FUNCTION_BLOCK basicValvulaCoester (* Logica do atuador Coester CSR (Modbus TCP) *)
  (* Standard: 61499-2 *)
  (* Version 2.5, 12/11/2026, Hidryco, Hidryco, 2.5: mapa revisado pelo MN_065 rev.3 (Modbus RTU, painel BLE): leitura 101-109 e comandos conferidos; posicao (word 105) = bits 0-7 parte inteira, bits 8-15 parte decimal - usa so o byte baixo, sem filtro de faixa (antes a word inteira dava valores acima de 1000). 2.4: posicao (Word 5) so atualiza com leitura de 0 a 100; fora da faixa mantem a ultima valida (antes era limitada, e um valor acima de 1000 virava 100 %%). 2.3: falha do atuador (alarmes da comunicacao) nao bloqueia o comando (fica disponivel em automatico) e nao muda a cor (sem animacao de falha); continua no alarme, no STS_ALARME e no diagnostico. 2.2: stsAlarme para a IO List da Nereda. 2.1: leituras 100 a 108 (posicao, torque, temperatura, tempo de percurso, status 2, alarmes), falha do atuador, posicionar por comando e parar so com cfgPosicionador (Word 2 de escrita). 2.0: refeito simples. *)
  PACKAGE Hidryco.HidrycoLib;
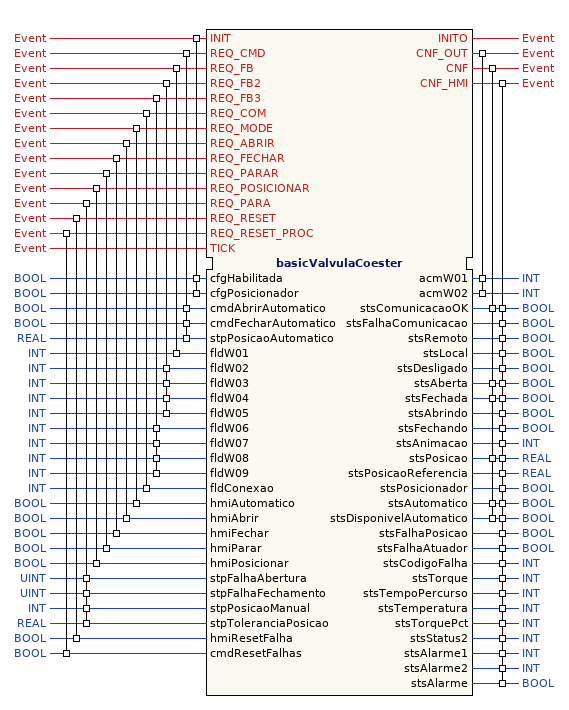
  EVENT_INPUT
    INIT WITH cfgHabilitada, cfgPosicionador; (* Inicializacao *)
    REQ_CMD WITH cmdAbrirAutomatico, cmdFecharAutomatico, stpPosicaoAutomatico; (* Processo: comandos do automatico *)
    REQ_FB WITH fldW01; (* Leitura Modbus: status 1 (endereco 100) *)
    REQ_FB2 WITH fldW02, fldW03, fldW04, fldW05; (* Leitura Modbus: enderecos 101 a 104 *)
    REQ_FB3 WITH fldW06, fldW07, fldW08, fldW09; (* Leitura Modbus: enderecos 105 a 108 *)
    REQ_COM WITH fldConexao; (* Status da conexao Modbus (connStatusInt) *)
    REQ_MODE WITH hmiAutomatico; (* IHM: modo *)
    REQ_ABRIR WITH hmiAbrir; (* IHM: abrir (manual) *)
    REQ_FECHAR WITH hmiFechar; (* IHM: fechar (manual) *)
    REQ_PARAR WITH hmiParar; (* IHM: parar (manual, so posicionador) *)
    REQ_POSICIONAR WITH hmiPosicionar; (* IHM: posicionar (manual, so posicionador) *)
    REQ_PARA WITH stpFalhaAbertura, stpFalhaFechamento, stpPosicaoManual, stpToleranciaPosicao; (* IHM: parametros *)
    REQ_RESET WITH hmiResetFalha; (* IHM: reset *)
    REQ_RESET_PROC WITH cmdResetFalhas; (* Processo: reset *)
    TICK; (* Base de tempo de 1 s *)
  END_EVENT
  EVENT_OUTPUT
    INITO; (* Inicializacao concluida *)
    CNF_OUT WITH acmW01, acmW02; (* Escrita Modbus (comando e posicao) *)
    CNF WITH stsDisponivelAutomatico, stsAberta, stsFechada, stsPosicao, stsAutomatico, stsComunicacaoOK; (* Status para o processo (na mudanca) *)
    CNF_HMI WITH stsComunicacaoOK, stsFalhaComunicacao, stsRemoto, stsLocal, stsDesligado, stsAberta, stsFechada, stsAbrindo, stsFechando, stsAnimacao, stsAutomatico, stsDisponivelAutomatico, stsFalhaPosicao, stsPosicionador, stsPosicao, stsPosicaoReferencia, stsFalhaAtuador, stsCodigoFalha, stsTorque, stsTempoPercurso, stsTemperatura, stsTorquePct, stsStatus2, stsAlarme1, stsAlarme2, stsAlarme; (* Status para a IHM (1 s e no comando) *)
  END_EVENT
  VAR_INPUT
    cfgHabilitada : BOOL := TRUE; (* FALSE = equipamento futuro: sem comunicacao esperada, sem alarme, fora do automatico *)
    cfgPosicionador : BOOL := FALSE; (* TRUE = posicionar e parar (700-VC-01); FALSE = so abrir e fechar *)
    cmdAbrirAutomatico : BOOL; (* Automatico: abrir *)
    cmdFecharAutomatico : BOOL; (* Automatico: fechar *)
    stpPosicaoAutomatico : REAL; (* Automatico: posicao desejada (%) - so posicionador *)
    fldW01 : INT; (* Word 1: status 1 (b0 local, b1 remoto, b2 desligado, b3 aberta, b4 fechada, b6 abrindo, b7 fechando) *)
    fldW02 : INT; (* Word 2: status 2 *)
    fldW03 : INT; (* Word 3: alarmes 1 *)
    fldW04 : INT; (* Word 4: alarmes 2 *)
    fldW05 : INT; (* Word 5: posicao (%) *)
    fldW06 : INT; (* Word 6: torque (Nm) *)
    fldW07 : INT; (* Word 7: tempo de percurso (s) *)
    fldW08 : INT; (* Word 8: temperatura (valor - 19 = graus C) *)
    fldW09 : INT; (* Word 9: torque (%) *)
    fldConexao : INT; (* Conexao Modbus: 1 = online *)
    hmiAutomatico : BOOL; (* IHM: TRUE = automatico *)
    hmiAbrir : BOOL; (* IHM: abrir *)
    hmiFechar : BOOL; (* IHM: fechar *)
    hmiParar : BOOL; (* IHM: parar *)
    hmiPosicionar : BOOL; (* IHM: posicionar *)
    stpFalhaAbertura : UINT; (* Tempo maximo para abrir (s); 0 = sem supervisao *)
    stpFalhaFechamento : UINT; (* Tempo maximo para fechar (s); 0 = sem supervisao *)
    stpPosicaoManual : INT; (* Posicao desejada em manual (%) *)
    stpToleranciaPosicao : REAL; (* Tolerancia da posicao (%); 0 = 2 % *)
    hmiResetFalha : BOOL; (* IHM: reset *)
    cmdResetFalhas : BOOL; (* Processo: reset (vale com TRUE) *)
  END_VAR
  VAR_OUTPUT
    acmW01 : INT; (* Word 1 de escrita (endereco 0): pulso b0 abrir, b1 fechar, b2 parar, b4 posicionar, b8 quitar alarmes *)
    acmW02 : INT; (* Word 2 de escrita (endereco 1): posicao desejada 0-100 % (so posicionador) *)
    stsComunicacaoOK : BOOL; (* Comunicacao OK *)
    stsFalhaComunicacao : BOOL; (* Falha de comunicacao *)
    stsRemoto : BOOL; (* Seletor em remoto *)
    stsLocal : BOOL; (* Seletor em local *)
    stsDesligado : BOOL; (* Seletor em desligado *)
    stsAberta : BOOL; (* Aberta *)
    stsFechada : BOOL; (* Fechada *)
    stsAbrindo : BOOL; (* Abrindo *)
    stsFechando : BOOL; (* Fechando *)
    stsAnimacao : INT; (* 0 fechada, 1 aberta, 2 falha, 3 intermediaria parada, 4 abrindo, 5 fechando *)
    stsPosicao : REAL; (* Posicao real (%) - Word 5 *)
    stsPosicaoReferencia : REAL; (* Ultima posicao enviada (%) *)
    stsPosicionador : BOOL; (* Copia de cfgPosicionador para a IHM *)
    stsAutomatico : BOOL; (* Modo automatico *)
    stsDisponivelAutomatico : BOOL; (* Pode ser comandada pelo automatico *)
    stsFalhaPosicao : BOOL; (* Nao abriu / nao fechou / nao posicionou no tempo (memorizada ate o reset) *)
    stsFalhaAtuador : BOOL; (* Falha do atuador (memorizada ate o reset) *)
    stsCodigoFalha : INT; (* Codigo da falha do atuador *)
    stsTorque : INT; (* Torque (Nm) *)
    stsTempoPercurso : INT; (* Tempo de percurso (s) *)
    stsTemperatura : INT; (* Temperatura (graus C) *)
    stsTorquePct : INT; (* Torque (%) *)
    stsStatus2 : INT; (* Word 2 *)
    stsAlarme1 : INT; (* Word 3 *)
    stsAlarme2 : INT; (* Word 4 *)
    stsAlarme : BOOL; (* Alarme: falha de comunicacao OU falha do atuador OU nao abriu/fechou/posicionou *)
  END_VAR
  VAR
    initDone : BOOL;
    comRecebido : BOOL;
    bComOk : BOOL;
    w01 : WORD;
    w02 : WORD;
    w03 : WORD;
    w04 : WORD;
    bFalhaAtiva : BOOL;
    codAtivo : INT;
    bAuto : BOOL := TRUE;
    bCmdMan : INT;
    bSpMan : REAL;
    bForca : BOOL;
    bPode : BOOL;
    bAlvo : INT;
    bAlvoAnt : INT := -1;
    bSp : REAL;
    bSpEnviado : REAL;
    bSubindo : BOOL;
    cBanda : REAL := 2.0;
    rTol : REAL;
    tLim : DINT;
    wPulso : WORD;
    tPulso : INT;
    cTempoPulso : INT := 2;
    wCmd : WORD;
    tReset : INT;
    tPos : INT;
    oldW01 : INT := -1;
    oldW02 : INT := -1;
    oldProc : INT := -1;
    oldPos : REAL := -1.0;
    nProc : INT;
    primeiro : BOOL := TRUE;
  END_VAR
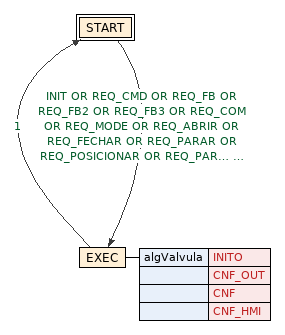
  EC_STATES
    START; (* Estado inicial *)
    EXEC : algValvula -> INITO, -> CNF_OUT, -> CNF, -> CNF_HMI; (* Executa a logica; o algoritmo decide quais eventos saem *)
  END_STATES
  EC_TRANSITIONS
    START TO EXEC := INIT OR REQ_CMD OR REQ_FB OR REQ_FB2 OR REQ_FB3 OR REQ_COM OR REQ_MODE OR REQ_ABRIR OR REQ_FECHAR OR REQ_PARAR OR REQ_POSICIONAR OR REQ_PARA OR REQ_RESET OR REQ_RESET_PROC OR TICK;
    EXEC TO START := 1;
  END_TRANSITIONS
  ALGORITHM algValvula IN ST: (* Logica completa da valvula (um unico algoritmo) *)
(* =====================================================================
   basicValvulaCoester 2.1 - logica do CAT Atuador_Coester (HidrycoLib)
   Atuador Coester CSR por Modbus TCP (mapa medido em campo):
   - leitura 100..108 = Words 1 a 9: status 1, status 2, alarmes 1 e 2,
     posicao (%), torque (Nm), tempo de percurso (s), temperatura (-19),
     torque (%);
   - escrita 0..1: Word 1 = comando EM PULSO de cTempoPulso s (b0 abrir,
     b1 fechar, b2 parar, b4 posicionar, b8 quitar alarmes); Word 2 =
     posicao desejada 0-100 %. O atuador retem o comando (MN_058 4.2.22);
     posicionar e "por comando" (padrao, MN_058 4.2.11): grava a Word 2 e
     pulsa o b4.
   - cfgPosicionador = TRUE (700-VC-01): posicionar e parar; no automatico
     segue stpPosicaoAutomatico e reposiciona quando ela muda cBanda (2 %)
     ou mais. FALSE: so abrir e fechar.
   - so comanda em remoto e com comunicacao OK; voltar a remoto repete o
     comando vigente; em manual cada botao repete o pulso;
   - "nao abriu / nao fechou / nao posicionou": o fim de curso (ou a
     posicao, com a tolerancia) nao veio no tempo configurado (0 = sem
     supervisao); memoriza ate o reset e pulsa parar;
   - falha do atuador: status 2 b0-b2, alarme 1 b1-b12, alarme 2 b0, b1,
     b4-b8; memoriza ate o reset; so informa (alarme e diagnostico):
     nao bloqueia o comando nem muda a cor da valvula;
   - cfgHabilitada = FALSE (equipamento futuro): sem alarme, fora do automatico.
   ===================================================================== *)

INITO   := FALSE;
CNF_OUT := FALSE;
CNF     := FALSE;
CNF_HMI := FALSE;

IF REQ_COM THEN
    comRecebido := TRUE;
END_IF;
IF INIT THEN
    initDone := TRUE;
    INITO    := TRUE;
END_IF;
IF NOT initDone THEN
    RETURN;
END_IF;

(* ---- 1. Leituras ---- *)
bComOk := cfgHabilitada AND comRecebido AND (fldConexao = 1);
w01 := INT_TO_WORD(fldW01);
w02 := INT_TO_WORD(fldW02);
w03 := INT_TO_WORD(fldW03);
w04 := INT_TO_WORD(fldW04);
IF bComOk THEN
    stsLocal     := (w01 AND 16#0001) <> 16#0000;
    stsRemoto    := (w01 AND 16#0002) <> 16#0000;
    stsDesligado := (w01 AND 16#0004) <> 16#0000;
    stsAberta    := (w01 AND 16#0008) <> 16#0000;
    stsFechada   := (w01 AND 16#0010) <> 16#0000;
    stsAbrindo   := (w01 AND 16#0040) <> 16#0000;
    stsFechando  := (w01 AND 16#0080) <> 16#0000;
    (* posicao (MN_065 rev.3, painel BLE, word 105): bits 0-7 = parte inteira (%), bits 8-15 = parte
       decimal; usa so o byte baixo (parte inteira) *)
    stsPosicao := INT_TO_REAL(WORD_TO_INT(INT_TO_WORD(fldW05) AND 16#00FF));
    stsTorque        := fldW06;
    stsTempoPercurso := fldW07;
    stsTemperatura   := fldW08 - 19;
    stsTorquePct     := fldW09;
    stsStatus2       := fldW02;
    stsAlarme1       := fldW03;
    stsAlarme2       := fldW04;
    bFalhaAtiva := ((w02 AND 16#0007) <> 16#0000) OR ((w03 AND 16#1FFE) <> 16#0000) OR ((w04 AND 16#01F3) <> 16#0000);
ELSE
    stsLocal := FALSE; stsRemoto := FALSE; stsDesligado := FALSE;
    stsAberta := FALSE; stsFechada := FALSE; stsAbrindo := FALSE; stsFechando := FALSE;
    bFalhaAtiva := FALSE;                      (* posicao e medicoes ficam no ultimo valor lido *)
END_IF;
stsComunicacaoOK    := bComOk;
stsFalhaComunicacao := cfgHabilitada AND NOT bComOk;
stsPosicionador     := cfgPosicionador;

(* codigo da falha ativa de maior prioridade (texto na IHM) *)
codAtivo := 0;
IF bFalhaAtiva THEN
    IF ((w02 AND 16#0001) <> 16#0000) OR ((w03 AND 16#0800) <> 16#0000) THEN codAtivo := 1;      (* falta de fase *)
    ELSIF ((w02 AND 16#0002) <> 16#0000) OR ((w03 AND 16#0040) <> 16#0000) THEN codAtivo := 2;   (* sobreaquecimento *)
    ELSIF ((w02 AND 16#0004) <> 16#0000) OR ((w03 AND 16#1000) <> 16#0000) THEN codAtivo := 3;   (* sem programacao *)
    ELSIF (w03 AND 16#0002) <> 16#0000 THEN codAtivo := 4;   (* parada local de emergencia *)
    ELSIF (w03 AND 16#0004) <> 16#0000 THEN codAtivo := 5;   (* torque na abertura *)
    ELSIF (w03 AND 16#0008) <> 16#0000 THEN codAtivo := 6;   (* torque no fechamento *)
    ELSIF (w03 AND 16#0010) <> 16#0000 THEN codAtivo := 7;   (* travado *)
    ELSIF (w03 AND 16#0020) <> 16#0000 THEN codAtivo := 8;   (* operacao incompleta *)
    ELSIF (w03 AND 16#0080) <> 16#0000 THEN codAtivo := 9;   (* falha ao energizar o motor *)
    ELSIF (w03 AND 16#0100) <> 16#0000 THEN codAtivo := 10;  (* motor energizado apos fim de curso *)
    ELSIF (w03 AND 16#0200) <> 16#0000 THEN codAtivo := 11;  (* motor energizado apos parada *)
    ELSIF (w03 AND 16#0400) <> 16#0000 THEN codAtivo := 12;  (* falha de comando *)
    ELSIF (w04 AND 16#0001) <> 16#0000 THEN codAtivo := 13;  (* tensao alta *)
    ELSIF (w04 AND 16#0002) <> 16#0000 THEN codAtivo := 14;  (* tensao baixa *)
    ELSIF (w04 AND 16#0030) <> 16#0000 THEN codAtivo := 15;  (* fim de curso mecanico ultrapassado *)
    ELSIF (w04 AND 16#00C0) <> 16#0000 THEN codAtivo := 16;  (* fim de curso programado ultrapassado *)
    ELSIF (w04 AND 16#0100) <> 16#0000 THEN codAtivo := 17;  (* cartao de rede nao detectado *)
    END_IF;
    stsFalhaAtuador := TRUE;                   (* memoriza ate o reset *)
    stsCodigoFalha  := codAtivo;
END_IF;

(* ---- 2. Reset (IHM ou processo) ---- *)
IF (REQ_RESET AND hmiResetFalha) OR (REQ_RESET_PROC AND cmdResetFalhas) THEN
    stsFalhaAtuador := bFalhaAtiva;            (* continua se a falha ainda esta ativa no atuador *)
    IF NOT bFalhaAtiva THEN
        stsCodigoFalha := 0;
    END_IF;
    stsFalhaPosicao := FALSE;
    tPos   := 0;
    tReset := 3;                               (* quitar alarmes no atuador por 3 s *)
END_IF;
IF TICK AND (tReset > 0) THEN
    tReset := tReset - 1;
END_IF;

(* ---- 3. Modo, parametros e comandos manuais ---- *)
IF REQ_MODE THEN
    bAuto := hmiAutomatico;
    bCmdMan := 0;                              (* troca de modo: nenhum comando manual *)
END_IF;
IF stpToleranciaPosicao > 0.0 THEN
    rTol := stpToleranciaPosicao;
ELSE
    rTol := 2.0;
END_IF;
bForca := FALSE;
IF NOT bAuto THEN
    IF REQ_ABRIR AND hmiAbrir THEN bCmdMan := 1; bForca := TRUE; END_IF;
    IF REQ_FECHAR AND hmiFechar THEN bCmdMan := 2; bForca := TRUE; END_IF;
    IF cfgPosicionador THEN
        IF REQ_PARAR AND hmiParar THEN bCmdMan := 4; bForca := TRUE; END_IF;
        IF REQ_POSICIONAR AND hmiPosicionar THEN
            bCmdMan := 3; bForca := TRUE;
            bSpMan := LIMIT(0.0, INT_TO_REAL(stpPosicaoManual), 100.0);
        END_IF;
    END_IF;
END_IF;

(* ---- 4. Comando desejado: 0 nenhum, 1 abrir, 2 fechar, 3 posicionar, 4 parar ---- *)
bPode := bComOk AND stsRemoto;
bSp := bSpEnviado;
IF NOT bPode THEN
    bAlvo := 0;                                (* fora de remoto ou sem comunicacao: nao comanda *)
ELSIF stsFalhaPosicao THEN
    bAlvo := 4;                                (* nao abriu / nao fechou / nao posicionou: para *)
ELSIF bAuto THEN
    IF cfgPosicionador THEN
        bAlvo := 3;
        bSp := LIMIT(0.0, stpPosicaoAutomatico, 100.0);
    ELSIF cmdAbrirAutomatico AND NOT cmdFecharAutomatico THEN
        bAlvo := 1;
    ELSIF cmdFecharAutomatico AND NOT cmdAbrirAutomatico THEN
        bAlvo := 2;
    ELSE
        bAlvo := 0;
    END_IF;
ELSE
    bAlvo := bCmdMan;
    IF bCmdMan = 3 THEN
        bSp := bSpMan;
    END_IF;
END_IF;

(* ---- 5. Pulso de comando ---- *)
IF TICK AND (tPulso > 0) THEN
    tPulso := tPulso - 1;
END_IF;
IF (bAlvo <> bAlvoAnt) OR (bForca AND bPode) OR ((bAlvo = 3) AND (ABS(bSp - bSpEnviado) >= cBanda)) THEN
    CASE bAlvo OF
        1: wPulso := 16#0001;
        2: wPulso := 16#0002;
        3: wPulso := 16#0010;
        4: wPulso := 16#0004;
    ELSE
        wPulso := 16#0000;
    END_CASE;
    IF bAlvo = 3 THEN
        bSubindo   := bSp >= stsPosicao;
        bSpEnviado := bSp;
    ELSIF bAlvo = 1 THEN
        bSpEnviado := 100.0;
    ELSIF bAlvo = 2 THEN
        bSpEnviado := 0.0;
    END_IF;
    IF wPulso <> 16#0000 THEN
        tPulso := cTempoPulso;
    ELSE
        tPulso := 0;
    END_IF;
    bAlvoAnt := bAlvo;
    tPos := 0;
END_IF;
IF tPulso > 0 THEN
    wCmd := wPulso;
ELSE
    wCmd := 16#0000;
END_IF;
IF tReset > 0 THEN
    wCmd := wCmd OR 16#0100;
END_IF;
acmW01 := WORD_TO_INT(wCmd);
acmW02 := REAL_TO_INT(LIMIT(0.0, bSpEnviado, 100.0));
stsPosicaoReferencia := bSpEnviado;
IF (acmW01 <> oldW01) OR (acmW02 <> oldW02) OR TICK OR primeiro THEN
    CNF_OUT := TRUE;
    oldW01 := acmW01;
    oldW02 := acmW02;
END_IF;

(* ---- 6. Nao abriu / nao fechou / nao posicionou ---- *)
IF TICK THEN
    tLim := 0;
    IF bPode THEN
        IF (bAlvo = 1) AND NOT stsAberta THEN
            tLim := UINT_TO_DINT(stpFalhaAbertura);
        ELSIF (bAlvo = 2) AND NOT stsFechada THEN
            tLim := UINT_TO_DINT(stpFalhaFechamento);
        ELSIF (bAlvo = 3) AND (ABS(stsPosicao - bSpEnviado) > rTol) THEN
            IF bSubindo THEN
                tLim := UINT_TO_DINT(stpFalhaAbertura);
            ELSE
                tLim := UINT_TO_DINT(stpFalhaFechamento);
            END_IF;
        END_IF;
    END_IF;
    IF tLim > 0 THEN
        tPos := tPos + 1;
        IF INT_TO_DINT(tPos) >= tLim THEN
            stsFalhaPosicao := TRUE;
        END_IF;
    ELSE
        tPos := 0;
    END_IF;
END_IF;

(* ---- 7. Saidas ---- *)
stsAutomatico := bAuto;
stsDisponivelAutomatico := bComOk AND stsRemoto AND bAuto AND NOT stsFalhaPosicao;   (* falha do atuador nao bloqueia *)
IF NOT bComOk OR stsFalhaPosicao THEN                                                (* falha do atuador nao muda a cor *)
    stsAnimacao := 2;
ELSIF stsAbrindo THEN
    stsAnimacao := 4;
ELSIF stsFechando THEN
    stsAnimacao := 5;
ELSIF stsAberta THEN
    stsAnimacao := 1;
ELSIF stsFechada THEN
    stsAnimacao := 0;
ELSE
    stsAnimacao := 3;
END_IF;
(* IO List da Nereda: alarme unico da valvula *)
stsAlarme := stsFalhaComunicacao OR stsFalhaAtuador OR stsFalhaPosicao;

(* ---- 8. Eventos: processo na mudanca (posicao a cada 1 %); IHM a cada 1 s e no comando ---- *)
nProc := BOOL_TO_INT(stsDisponivelAutomatico) + 2 * BOOL_TO_INT(stsAberta) + 4 * BOOL_TO_INT(stsFechada) +
         8 * BOOL_TO_INT(stsAutomatico) + 16 * BOOL_TO_INT(bComOk);
IF primeiro OR (nProc <> oldProc) OR (ABS(stsPosicao - oldPos) >= 1.0) THEN
    CNF := TRUE;
    oldProc := nProc;
    oldPos := stsPosicao;
END_IF;
IF primeiro OR TICK OR REQ_MODE OR REQ_ABRIR OR REQ_FECHAR OR REQ_PARAR OR REQ_POSICIONAR OR REQ_PARA OR REQ_RESET OR REQ_RESET_PROC OR
   REQ_FB OR REQ_COM THEN
    CNF_HMI := TRUE;
END_IF;
primeiro := FALSE;
  END_ALGORITHM
END_FUNCTION_BLOCK
